(* IEC 61131-3 sources: PortalRobot/Portal_robot/Device/application/ST/ST_MAGAZINE, 26 files *)

(* ---- E_MAGAZINE_OPERATION.st ---- *)
{attribute 'qualified_only'}
{attribute 'strict'}
TYPE E_MAGAZINE_OPERATION :
(
	NONE         := 0,
	PUT          := 1,
	TAKE         := 2,
	CHANGE       := 3,
	RETURN_BLANK := 4
);
END_TYPE

(* ---- E_MAGAZINE_STATE.st ---- *)
{attribute 'qualified_only'}
{attribute 'strict'}
TYPE E_MAGAZINE_STATE :
(
	DISABLED,
	IDLE,
	CHOOSE,
	PREPARE_STEP,
	ROBOT_COMMAND,
	RELEASE_ROBOT_COMMAND,
	NEXT,
	DONE,
	ERROR
);
END_TYPE

(* ---- E_TWO_PALLET_STATE.st ---- *)
{attribute 'qualified_only'}
{attribute 'strict'}
TYPE E_TWO_PALLET_STATE :
(
	IDLE := 0,
	AUTO_LOWER := 20,
	AUTO_MOVE_TO_EXCHANGE := 30,
	AUTO_SELECT_PALLET := 40,
	AUTO_MOVE_TO_WORK := 50,
	AUTO_RAISE := 60,
	MANUAL_LOWER := 100,
	MANUAL_RAISE := 110,
	MANUAL_SELECT_PALLET := 120,
	MANUAL_MOVE := 130,
	MANUAL_HOME := 150,
	MANUAL_JOG := 160,
	MANUAL_LOCK := 170,
	MANUAL_STOP := 180
);
END_TYPE

(* ---- ST_MAGAZINE_CALIBRATION.st ---- *)
TYPE ST_MAGAZINE_CALIBRATION :
STRUCT
	uiMethod : UINT := UINT#1; // 1: база и мировые X/Y; 3: база A и направления B/C
	astReference : ARRAY [1..2] OF ST_POINT; // B: последний слот первого ряда; C: первый слот последнего ряда
END_STRUCT
END_TYPE

(* ---- ST_MAGAZINE_CALIBRATION_STATUS.st ---- *)
TYPE ST_MAGAZINE_CALIBRATION_STATUS :
STRUCT
	uiMethod : UINT := UINT#1;
	xChangeAllowed : BOOL;
	xCaptureAllowed : BOOL;
	xSaveAllowed : BOOL;
	xReferenceCaptureAllowed : BOOL;
	xReferenceSaveAllowed : BOOL;
	xMoveAAllowed : BOOL;
	xMoveBAllowed : BOOL;
	xMoveCAllowed : BOOL;
	xReady : BOOL;
	uiReason : UINT;
	astPoints : ARRAY [1..3] OF ST_POINT; // Согласованная публикация A/B/C вместе с методом для экспорта
END_STRUCT
END_TYPE

(* ---- ST_MAGAZINE_COMMAND.st ---- *)
TYPE ST_MAGAZINE_COMMAND :
STRUCT
	xEnable  : BOOL; // Импульс включения магазина
	xDisable : BOOL; // Импульс отключения магазина
	xExecute : BOOL; // Запуск выбранной операции
	xStop    : BOOL; // Остановка текущей операции
	eOperation : E_MAGAZINE_OPERATION; // Операция автоматического цикла
	iTakeSlot  : SINT; // Слот заготовки для TAKE/CHANGE
	iPutSlot   : SINT; // Слот укладки для PUT/CHANGE/RETURN_BLANK
END_STRUCT
END_TYPE

(* ---- ST_MAGAZINE_DIAG.st ---- *)
TYPE ST_MAGAZINE_DIAG :
STRUCT
	eState : E_MAGAZINE_STATE := E_MAGAZINE_STATE.DISABLED; // Текущее состояние автомата магазина
	stWarning : ST_WARNING_EVENT; // Последнее предупреждение магазина
END_STRUCT
END_TYPE

(* ---- ST_MAGAZINE_ERROR.st ---- *)
TYPE ST_MAGAZINE_ERROR :
STRUCT
	WRONG_OPERATION : BOOL; // Операция не может быть выбрана
	NO_BLANK        : BOOL; // В магазине нет доступной заготовки
	NO_FREE_SLOT    : BOOL; // В магазине нет свободного слота
	INVALID_SLOT    : BOOL; // Номер слота находится вне матрицы
	SLOT_CONTENT    : BOOL; // Содержимое выбранного слота не соответствует операции
	ROBOT_ERROR     : BOOL; // Робот завершил команду с ошибкой
	GLOBAL_STOP     : BOOL; // Получена глобальная ошибка ячейки
	GEOMETRY_ERROR  : BOOL; // Геометрия магазина задана неверно
END_STRUCT
END_TYPE

(* ---- ST_MAGAZINE_ERRORS.st ---- *)
TYPE ST_MAGAZINE_ERRORS :
STRUCT
	dwErrorActive : DWORD; // Битовая маска активных ошибок
	dwErrorLast   : DWORD; // Битовая маска последних ошибок
	dwAlarmActive : DWORD; // Собственные аварии магазина для общего журнала
	stErrorActive : ST_MAGAZINE_ERROR; // Расшифровка активных ошибок
	stErrorLast   : ST_MAGAZINE_ERROR; // Расшифровка последних ошибок
END_STRUCT
END_TYPE

(* ---- ST_MAGAZINE_FAULT_REQUEST.st ---- *)
TYPE ST_MAGAZINE_FAULT_REQUEST :
STRUCT
	xEnabled        : BOOL; // Глобальное разрешение диагностической инъекции
	xWrongOperation : BOOL; // Импульс недопустимой операции
	xNoBlank        : BOOL; // Импульс отсутствия заготовки
	xNoFreeSlot     : BOOL; // Импульс отсутствия свободного слота
	xInvalidSlot    : BOOL; // Импульс недопустимого номера слота
	xSlotContent    : BOOL; // Импульс несоответствия содержимого слота
	xGeometry       : BOOL; // Импульс недопустимой геометрии магазина
END_STRUCT
END_TYPE

(* ---- ST_MAGAZINE_FRAME.st ---- *)
TYPE ST_MAGAZINE_FRAME :
STRUCT
	stAxisX : ST_MAGAZINE_VECTOR;
	stAxisY : ST_MAGAZINE_VECTOR;
	stAxisZ : ST_MAGAZINE_VECTOR;
	xReady : BOOL;
	uiReason : UINT; // 0 готово; 1 нет базы/Z; 2 неверный метод/сетка; 3 нет B/C; 4 вырожденная плоскость; 5 внешний робот
END_STRUCT
END_TYPE

(* ---- ST_MAGAZINE_HMI_COMMAND.st ---- *)
TYPE ST_MAGAZINE_HMI_COMMAND :
STRUCT
	{attribute 'symbol' := 'read'}
	xEnable : BOOL; // Импульс включения технологической логики магазина
	{attribute 'symbol' := 'read'}
	xDisable : BOOL; // Импульс отключения технологической логики магазина
	{attribute 'symbol' := 'read'}
	xStop : BOOL; // Остановить выполняемую операцию магазина
	{attribute 'symbol' := 'read'}
	xReset : BOOL; // Сброс ошибок магазина
	{attribute 'symbol' := 'read'}
	xFill : BOOL; // Заполнить кассету заготовками по текущей карте типов
	{attribute 'symbol' := 'read'}
	xClear : BOOL; // Полностью очистить кассету
	xCycleSlot : BOOL; // Переключить содержимое выбранного слота
	{attribute 'symbol' := 'read'}
	xApplySlot : BOOL; // Явно записать состояние и тип выбранного слота
	{attribute 'symbol' := 'read'}
	xApplyPitchX : BOOL; // Применить новый шаг слотов по X
	{attribute 'symbol' := 'read'}
	xApplyPitchY : BOOL; // Применить новый шаг слотов по Y
	uiEditSlot : UINT; // Слот кассеты, 1..120
	uiEditDetailType : UINT; // 0=NONE, 1=BLANK, 2=DETAIL
	uiEditProductType : UINT; // Тип изделия 1..3; для NONE игнорируется
	lrEditPitchX : LREAL; // Запрошенный шаг слотов по X
	lrEditPitchY : LREAL; // Запрошенный шаг слотов по Y
END_STRUCT
END_TYPE

(* ---- ST_MAGAZINE_INVENTORY.st ---- *)
TYPE ST_MAGAZINE_INVENTORY :
STRUCT
	aSlots : ARRAY [1..GVL_CELL_SETTINGS.MagazineSlots] OF ST_DETAIL; // Единственная статичная кассета
END_STRUCT
END_TYPE

(* ---- ST_MAGAZINE_STATUS.st ---- *)
TYPE ST_MAGAZINE_STATUS :
STRUCT
	xEnabled         : BOOL; // Магазин включен в работу
	xDisablePending  : BOOL; // Отключение выполнится после выхода робота и завершения операции
	xPowerAllowed    : BOOL; // Команда включения/отключения может быть принята
	xEnableSequenceAllowed : BOOL; // PLC разрешает ввести подготовленный магазин в автомат
	xEnableCheckRobotReady : BOOL; // Диагностика готовности роботной операции; не блокирует включение
	xEnableCheckRobotReleased : BOOL; // Диагностика положения робота; не блокирует включение
	xEnableCheckNoError : BOOL; // Нет ошибок магазина и глобальных ошибок ячейки
	xEnableCheckContent : BOOL; // Содержимое кассеты допускает полезную операцию
	xEnableCheckGeometry : BOOL; // Матрица содержит от 1 до 120 активных слотов
	xFillAllowed     : BOOL; // Кнопка заполнения магазина заготовками доступна
	xClearAllowed    : BOOL; // Кнопка очистки магазина доступна
	xEditAllowed     : BOOL; // Содержимое разрешено менять только у выключенного магазина
	xPitchEditAllowed : BOOL; // Общий шаг X/Y можно менять только при выключенных обоих магазинах
	xReady 			 : BOOL; // Магазин готов принять команду
	xBusy  			 : BOOL; // Выполняется операция магазина
	xDone  			 : BOOL; // Операция магазина завершена
	xError          : BOOL; // Магазин находится в ошибке
	xRobotStopRequired : BOOL; // Ошибка магазина требует зависимой аварии робота
	xOutBlank        : BOOL; // В магазине не осталось свободных заготовок
	xOutFreeSlot     : BOOL; // В магазине не осталось свободных слотов
	xCanTake         : BOOL; // Операция TAKE доступна по содержимому магазина
	xCanPut          : BOOL; // Операция PUT доступна по содержимому магазина
	xCanChange       : BOOL; // Операция CHANGE доступна по содержимому магазина
	xCanEnable       : BOOL; // Содержимое позволяет взять/положить груз; не блокирует включение
	xFinished        : BOOL; // Палета завершена; защёлка до смены/правки её рабочего содержимого
	udiProducedPartsTotal : UDINT; // Подтверждённые укладки готовой детали с момента запуска PLC
	uiMagazineId    : UINT; // 1 или 2
	iCurrentBlank    : SINT; // Минимальный номер заготовки в матрице
	iCurrentFreeSlot : SINT; // Минимальный номер свободного слота в матрице
	iSelectedBlank   : SINT; // Номер заготовки, выбранной для текущей операции
	iSelectedFreeSlot: SINT; // Номер свободного слота, выбранного для текущей операции
	eGrantedOperation: E_MAGAZINE_OPERATION; // Доступная операция по текущему состоянию магазина
	eActualOperation : E_MAGAZINE_OPERATION; // Выполняемая операция магазина
	stTypeStatus     : ST_MAGAZINE_TYPE_STATUS; // Содержимое кассеты по типам
END_STRUCT
END_TYPE

(* ---- ST_MAGAZINE_TYPE_STATUS.st ---- *)
TYPE ST_MAGAZINE_TYPE_STATUS :
STRUCT
	aiBlankSlot    : ARRAY [1..3] OF SINT; // Первая заготовка каждого типа
	aiFreeSlot     : ARRAY [1..3] OF SINT; // Первый свободный слот каждого типа
	auiBlankCount  : ARRAY [1..3] OF UINT; // Количество заготовок каждого типа
	auiDetailCount : ARRAY [1..3] OF UINT; // Количество готовых деталей каждого типа
	auiFreeCount   : ARRAY [1..3] OF UINT; // Количество свободных слотов каждого типа
END_STRUCT
END_TYPE

(* ---- ST_MAGAZINE_VECTOR.st ---- *)
TYPE ST_MAGAZINE_VECTOR :
STRUCT
	X : LREAL;
	Y : LREAL;
	Z : LREAL;
END_STRUCT
END_TYPE

(* ---- ST_TWO_PALLET_COMMAND.st ---- *)
TYPE ST_TWO_PALLET_COMMAND :
STRUCT
	xEnable : BOOL;
	xConfirm : BOOL;
	xStart : BOOL; // Атомарно подтвердить актуальную расстановку и включить магазин
	xRejectStart : BOOL; // Оператор ответил «Нет» в предпусковом окне
	xDisable : BOOL;
	xSwap : BOOL;
	xPowerOn : BOOL;
	xPowerOff : BOOL;
	xDriveReset : BOOL;
	xHome : BOOL;
	xLower : BOOL;
	xRaise : BOOL;
	xSelectPallet : BOOL;
	xLockIn : BOOL;
	xLockOut : BOOL;
	xStopIn : BOOL;
	xStopOut : BOOL;
	xMoveToExchange : BOOL;
	xMoveToWork : BOOL;
	xStop : BOOL;
	xReset : BOOL;
	xJogPositive : BOOL;
	xJogNegative : BOOL;
	xJogRelease : BOOL;
	xTeachOperator : BOOL; // Запомнить текущую координату переключения/операторской зоны
	xTeachWork : BOOL; // Запомнить текущую рабочую координату выбранной палеты у робота
	uiPallet : UINT; // Номер подтверждаемой/выбираемой палеты, 1..2
	udiRevision : UDINT; // Ревизия расстановки для команды подтверждения
END_STRUCT
END_TYPE

(* ---- ST_TWO_PALLET_CONFIG.st ---- *)
TYPE ST_TWO_PALLET_CONFIG :
STRUCT
	xConfigured : BOOL; // Не выставляется автоматически; параметры проверены на механизме
	xP1LockOut : BOOL; // Legacy: используется только при переносе старой RETAIN-конфигурации
	lrExchange : LREAL;
	lrWorkP1 : LREAL;
	lrWorkP2 : LREAL;
	lrHome : LREAL;
	lrTolerance : LREAL;
	lrVelocity : LREAL;
	lrAcceleration : LREAL;
	lrDeceleration : LREAL;
	lrJerk : LREAL;
	tCylinder : TIME;
	tMove : TIME;
	tHome : TIME;
	tPulse : TIME;
	xSignalPatternsConfigured : BOOL;
	uiP1Signals : UINT; // Биты 0..5: LiftDown, LiftUp, LockIn, LockOut, StopIn, StopOut
	uiP2Signals : UINT; // Полные ожидаемые состояния шести герконов для П2 у робота
END_STRUCT
END_TYPE

(* ---- ST_TWO_PALLET_DIAG.st ---- *)
TYPE ST_TWO_PALLET_DIAG :
STRUCT
	eState : E_TWO_PALLET_STATE := E_TWO_PALLET_STATE.IDLE;
	eFaultState : E_TWO_PALLET_STATE := E_TWO_PALLET_STATE.IDLE;
	uiReason : UINT; // Первая причина блокировки подтверждения/включения магазина
	stWarning : ST_WARNING_EVENT;
END_STRUCT
END_TYPE

(* ---- ST_TWO_PALLET_ERROR.st ---- *)
TYPE ST_TWO_PALLET_ERROR :
STRUCT
	DRIVE_ERROR : BOOL;
	SENSOR_CONTRADICTION : BOOL;
	CYLINDER_TIMEOUT : BOOL;
	MOTION_TIMEOUT : BOOL;
	LOGIC_ERROR : BOOL;
	SEQUENCE_INTERRUPTED : BOOL;
END_STRUCT
END_TYPE

(* ---- ST_TWO_PALLET_ERRORS.st ---- *)
TYPE ST_TWO_PALLET_ERRORS :
STRUCT
	dwErrorActive : DWORD;
	dwErrorLast : DWORD;
	dwAlarmActive : DWORD;
	stErrorActive : ST_TWO_PALLET_ERROR;
	stErrorLast : ST_TWO_PALLET_ERROR;
END_STRUCT
END_TYPE

(* ---- ST_TWO_PALLET_INPUT.st ---- *)
TYPE ST_TWO_PALLET_INPUT :
STRUCT
	xIoMapped : BOOL; // Подтверждается наладчиком после привязки и проверки физических I/O
	xLiftDown : BOOL;
	xLiftUp : BOOL;
	xLockIn : BOOL;
	xLockOut : BOOL;
	xStopIn : BOOL;
	xStopOut : BOOL;
	xLimitNegative : BOOL;
	xLimitPositive : BOOL;
	xHomeSensor : BOOL; // Только датчик каретки, не палет
	xAxisBound : BOOL;
	xPowered : BOOL;
	xHomed : BOOL;
	xStandstill : BOOL;
	xDriveError : BOOL;
	xMotionDone : BOOL;
	lrPosition : LREAL;
END_STRUCT
END_TYPE

(* ---- ST_TWO_PALLET_OUTPUT.st ---- *)
TYPE ST_TWO_PALLET_OUTPUT :
STRUCT
	xLiftUp : BOOL;
	xLiftDown : BOOL;
	xLockOut : BOOL;
	xLockIn : BOOL;
	xStopOut : BOOL;
	xStopIn : BOOL;
	xPowerOn : BOOL;
	xPowerOff : BOOL;
	xDriveReset : BOOL;
	xHome : BOOL;
	xMove : BOOL;
	xStop : BOOL;
	xJogPositive : BOOL;
	xJogNegative : BOOL;
	xTeachOperator : BOOL;
	xTeachWork : BOOL;
	lrTarget : LREAL;
END_STRUCT
END_TYPE

(* ---- ST_TWO_PALLET_REQUEST.st ---- *)
TYPE ST_TWO_PALLET_REQUEST :
STRUCT
	uiMagazine : UINT; // 0: конфигурация линии; 1..2: отдельный магазин
	uiCommand : UINT;
	uiValue : UINT;
	uiSlot : UINT;
	uiContent : UINT;
	uiProductType : UINT;
	udiRevision : UDINT;
	Config : ST_TWO_PALLET_CONFIG;
END_STRUCT
END_TYPE

(* ---- ST_TWO_PALLET_STATUS.st ---- *)
TYPE ST_TWO_PALLET_STATUS :
STRUCT
	uiStep : UINT;
	uiFaultStep : UINT; // Шаг, на котором появился последний новый аварийный бит
	uiCandidate : UINT; // Расстановка, совместимая с датчиками; не измерение палет
	uiRobotPallet : UINT := 1; // Учётный номер, меняется только после подтверждения/завершения обмена
	uiSelected : UINT;
	udiRevision : UDINT;
	xEnabled : BOOL;
	xConfirmed : BOOL;
	xReady : BOOL;
	xBusy : BOOL;
	xError : BOOL;
	xHomeRequired : BOOL;
	xConfigValid : BOOL;
	xConfirmAllowed : BOOL;
	xStartAllowed : BOOL;
	xEnableAllowed : BOOL;
	xSwapAllowed : BOOL;
	xPowerAllowed : BOOL;
	xDriveResetAllowed : BOOL;
	xHomeAllowed : BOOL;
	xLowerAllowed : BOOL;
	xRaiseAllowed : BOOL;
	xSelectAllowed : BOOL;
	xLockAllowed : BOOL;
	xStopAllowed : BOOL;
	xMoveAllowed : BOOL;
	xJogAllowed : BOOL;
	xTeachOperatorAllowed : BOOL;
	xTeachWorkAllowed : BOOL;
	xResetAllowed : BOOL;
	xEditAllowed : BOOL;
	xEdit1Allowed : BOOL;
	xEdit2Allowed : BOOL;
	xLoadAllowed : BOOL; // Подтвердить загрузку текущей операторской палеты
	xConfigAllowed : BOOL;
	xCompleted : BOOL;
	xCommandAccepted : BOOL;
	uiReason : UINT;
	dwError : DWORD;
	stWarning : ST_WARNING_EVENT;
	Input : ST_TWO_PALLET_INPUT;
	rP1 : REAL; // Оценка нормализованного положения для 3D, не датчик палеты
	rP2 : REAL;
	rLift : REAL;
	xAutoSwapEnabled : BOOL; // Настройка автоматической смены палет
END_STRUCT
END_TYPE

(* ---- ST_TWO_PALLET_STORE.st ---- *)
TYPE ST_TWO_PALLET_STORE :
STRUCT
	astPallet : ARRAY [1..2] OF ST_MAGAZINE_INVENTORY;
	axLoaded : ARRAY [1..2] OF BOOL; // Снимается после обмена и каждого редактирования
END_STRUCT
END_TYPE
